(* IEC 61131-3 sources: SemantiST/benchmarks/defects/designed/d08_pin_lockout/buggy, 1 file *)

(* ---- target.st ---- *)
FUNCTION_BLOCK D08_PIN_LOCKOUT
VAR_INPUT
    Enter : BOOL;
    Code : INT;
END_VAR
VAR_OUTPUT
    Unlocked : BOOL;
    Locked : BOOL;
END_VAR
VAR
    lockTimer : TON;
    failures : INT;
    attempts : ARRAY[0..3] OF INT;
    lastEnter : BOOL;
END_VAR

lockTimer(IN := Locked, PT := T#500ms);
IF lockTimer.Q THEN
    (* defect: failures is not reset when the lock expires *)
    Locked := FALSE;
END_IF;
IF Enter AND NOT lastEnter AND NOT Locked THEN
    IF Code = 4711 THEN
        Unlocked := TRUE;
        failures := 0;
    ELSE
        Unlocked := FALSE;
        attempts[failures] := Code;
        failures := failures + 1;
        IF failures >= 3 THEN
            Locked := TRUE;
        END_IF;
    END_IF;
END_IF;
lastEnter := Enter;
END_FUNCTION_BLOCK
